(* IEC 61131-3 sources: llm-plc-st-eval/data/definitivo/claude-sonnet-4-6/B1/few_shot, 3 files *)

(* ---- ejec_1.st ---- *)
```st
FUNCTION_BLOCK FB_Motor
VAR_INPUT
    btnMarcha : BOOL; (* Boton de marcha *)
    btnParo   : BOOL; (* Boton de paro *)
    btnEmerg  : BOOL; (* Boton de paro de emergencia *)
END_VAR
VAR_OUTPUT
    motorOn : BOOL; (* Salida del motor *)
END_VAR
VAR
    bloqEmerg : BOOL; (* Bloqueo activo tras paro de emergencia *)
END_VAR

(* Si se activa emergencia: apagar motor y activar bloqueo *)
IF btnEmerg THEN
    bloqEmerg := TRUE;
    motorOn   := FALSE;

(* Si se pulsa paro: apagar motor (sin bloqueo) *)
ELSIF btnParo THEN
    motorOn := FALSE;

(* Arranque solo si no hay bloqueo de emergencia *)
ELSIF btnMarcha AND NOT bloqEmerg THEN
    motorOn := TRUE;
END_IF;

(* El bloqueo de emergencia se libera unicamente cuando
   btnEmerg ya no esta activo Y btnMarcha no esta pulsado,
   evitando rearranque involuntario al liberar el bloqueo *)
IF bloqEmerg AND NOT btnEmerg AND NOT btnMarcha THEN
    bloqEmerg := FALSE;
END_IF;

END_FUNCTION_BLOCK
```

(* ---- ejec_2.st ---- *)
```st
FUNCTION_BLOCK FB_Motor
VAR_INPUT
    btnMarcha : BOOL; (* Boton de marcha *)
    btnParo   : BOOL; (* Boton de paro *)
    btnEmerg  : BOOL; (* Boton de paro de emergencia *)
END_VAR
VAR_OUTPUT
    motorOn : BOOL; (* Salida del motor *)
END_VAR
VAR
    bloqEmerg : BOOL; (* Bloqueo activo tras emergencia *)
END_VAR

(* Activar bloqueo de emergencia; solo se libera al ciclo siguiente sin emergencia *)
IF btnEmerg THEN
    bloqEmerg := TRUE;
END_IF;

(* Logica de arranque/paro con autoretencion *)
(* Paro normal o emergencia detienen el motor                *)
(* El bloqueo impide rearranque hasta que se libere          *)
IF btnParo OR btnEmerg THEN
    motorOn := FALSE;
ELSIF btnMarcha AND NOT bloqEmerg THEN
    motorOn := TRUE;
END_IF;

(* Liberar bloqueo de emergencia solo cuando no hay emergencia ni motor en marcha *)
IF NOT btnEmerg AND NOT motorOn THEN
    bloqEmerg := FALSE;
END_IF;

END_FUNCTION_BLOCK
```

(* ---- ejec_3.st ---- *)
```st
FUNCTION_BLOCK FB_Motor
VAR_INPUT
    btnMarcha : BOOL; (* Boton de marcha *)
    btnParo   : BOOL; (* Boton de paro *)
    btnEmerg  : BOOL; (* Boton de paro de emergencia *)
END_VAR
VAR_OUTPUT
    motorOn : BOOL; (* Salida del contactor del motor *)
END_VAR
VAR
    bloqEmerg : BOOL; (* Bloqueo activo tras paro de emergencia *)
END_VAR

(* Activar bloqueo ante paro de emergencia; se mantiene hasta nuevo ciclo de paro normal *)
IF btnEmerg THEN
    bloqEmerg := TRUE;
END_IF;

(* Desbloquear solo cuando se pulsa paro sin emergencia activa *)
IF btnParo AND NOT btnEmerg THEN
    bloqEmerg := FALSE;
END_IF;

(* Logica de arranque con autoretencion:
   - Arranca si btnMarcha y no hay bloqueo de emergencia
   - Para si btnParo o btnEmerg                          *)
IF (btnParo OR btnEmerg) THEN
    motorOn := FALSE;
ELSIF btnMarcha AND NOT bloqEmerg THEN
    motorOn := TRUE;
END_IF;
(* Si ninguna condicion se cumple, motorOn conserva su estado anterior (autoretencion) *)

END_FUNCTION_BLOCK
```
